// Forçages actifs (docs/12 § 7), persistants
{attribute 'pack_mode' := '1'}
TYPE ST_MachineForce :
STRUCT
    eDeclared : E_DeclaredState;
    bStartBlocked : BOOL;
    nReason : USINT;
    tSince : LINT;
    tUntil : LINT;
    sBy : STRING(24);
    aStation : ARRAY[1..GVL_Const.MAX_STATIONS] OF ST_StationForce;
    aMover : ARRAY[1..GVL_Const.MAX_MOVERS] OF ST_MoverForce;
END_STRUCT
END_TYPE

(* stored: Version 1.1.0.1, ProductVersion 3.1.4024.12
   DUT ST_MachineForce: Id {73ee7676-d138-554d-b0e6-ddc340c3a649} *)
